// TIA Portal project "Yapisal Programlama" (V18)

(* hardware
DEVICE "S7-1200 station_1"  S7-1200 Station
   slot 0: "Rack_0"  S7-1200 Rack  Rack  V1.0
   slot 1: "PLC_1"  CPU 1214C DC/DC/Rly  6ES7 214-1HG40-0XB0  V4.6
*)

// ===== PLC "PLC_1"  CPU 1214C DC/DC/Rly =====

VAR_GLOBAL   // PLC tag table "Default tag table"
   "Start Butonu" AT %I0.0 : Bool;
   "Acil Stop Butonu" AT %I0.1 : Bool;
   "Reset Butonu" AT %I0.2 : Bool;
   "Yukarı Sensörü" AT %I0.3 : Bool;
   "Aşağı Sensörü" AT %I0.4 : Bool;
   "Piston Yukarı" AT %Q0.0 : Bool;
   "Piston Aşağı" AT %Q0.1 : Bool;
   "Sistem Start Mem" AT %M10.0 : Bool;
END_VAR

// folder: System blocks/Program resources

DATA_BLOCK "Counter 1"   // DB1
{ S7_Optimized_Access := 'TRUE' }
AUTHOR : Simatic
FAMILY : IEC
NAME : CNTR
VERSION : 1.0
// stored: InstanceOfName IEC_COUNTER
"IEC_COUNTER"
BEGIN
END_DATA_BLOCK

DATA_BLOCK "TIMER -1"   // DB2
{ S7_Optimized_Access := 'TRUE' }
AUTHOR : Simatic
FAMILY : IEC
NAME : IEC_TMR
VERSION : 1.0
// stored: InstanceOfName IEC_TIMER
"IEC_TIMER"
BEGIN
END_DATA_BLOCK

// folder: (top level)

FUNCTION "Normal Calisma" : Void   // FC1, LAD
{ S7_Optimized_Access := 'TRUE' }
VERSION : 0.1
BEGIN

REGION Network 1: SİSTEMİN BAŞLATILMASI
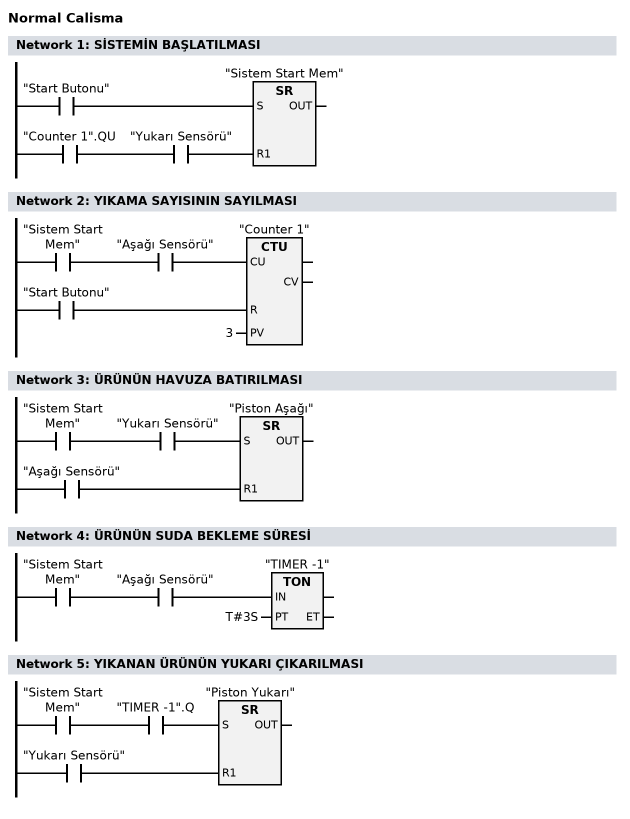
   RUNG wire#powerrail
      Contact( "Start Butonu" )
      S_SR(operand := "Sistem Start Mem", r1 := wire#w1)
   END_RUNG
   RUNG wire#powerrail
      Contact( "Counter 1".QU )
      Contact( "Yukarı Sensörü" )
   END_RUNG wire#w1
   // the same network as SCL:
   IF "Start Butonu" THEN
       "Sistem Start Mem" := TRUE;   // SR flip-flop
   END_IF;
   IF "Counter 1".QU AND "Yukarı Sensörü" THEN "Sistem Start Mem" := FALSE; END_IF;
END_REGION

REGION Network 2: YIKAMA SAYISININ SAYILMASI
   "Counter 1".CTU(CU := "Sistem Start Mem" AND "Aşağı Sensörü", R := "Start Butonu", PV := 3);
END_REGION

REGION Network 3: ÜRÜNÜN HAVUZA BATIRILMASI
   RUNG wire#powerrail
      Contact( "Sistem Start Mem" )
      Contact( "Yukarı Sensörü" )
      S_SR(operand := "Piston Aşağı", r1 := wire#w1)
   END_RUNG
   RUNG wire#powerrail
      Contact( "Aşağı Sensörü" )
   END_RUNG wire#w1
   // the same network as SCL:
   IF "Sistem Start Mem" AND "Yukarı Sensörü" THEN
       "Piston Aşağı" := TRUE;   // SR flip-flop
   END_IF;
   IF "Aşağı Sensörü" THEN "Piston Aşağı" := FALSE; END_IF;
END_REGION

REGION Network 4: ÜRÜNÜN SUDA BEKLEME SÜRESİ
   "TIMER -1".TON(IN := "Sistem Start Mem" AND "Aşağı Sensörü", PT := T#3S);
END_REGION

REGION Network 5: YIKANAN ÜRÜNÜN YUKARI ÇIKARILMASI
   RUNG wire#powerrail
      Contact( "Sistem Start Mem" )
      Contact( "TIMER -1".Q )
      S_SR(operand := "Piston Yukarı", r1 := wire#w1)
   END_RUNG
   RUNG wire#powerrail
      Contact( "Yukarı Sensörü" )
   END_RUNG wire#w1
   // the same network as SCL:
   IF "Sistem Start Mem" AND "TIMER -1".Q THEN
       "Piston Yukarı" := TRUE;   // SR flip-flop
   END_IF;
   IF "Yukarı Sensörü" THEN "Piston Yukarı" := FALSE; END_IF;
END_REGION
END_FUNCTION

FUNCTION "Acil Stop Calisma" : Void   // FC2, LAD
{ S7_Optimized_Access := 'TRUE' }
VERSION : 0.1
BEGIN

REGION Network 1: ACİL STOP BUTONUNA BASILDIĞINDA SİSTEMİN DURDURULMASI
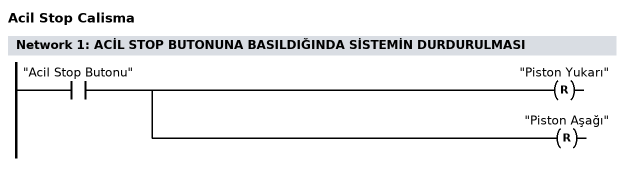
   RUNG wire#powerrail
      Contact( "Acil Stop Butonu" )
      wire#w1
      R_Coil( "Piston Yukarı" )
   END_RUNG
   RUNG wire#w1
      R_Coil( "Piston Aşağı" )
   END_RUNG
   // the same network as SCL:
   IF "Acil Stop Butonu" THEN
       "Piston Yukarı" := FALSE;
       "Piston Aşağı" := FALSE;
   END_IF;
END_REGION
END_FUNCTION

FUNCTION "Reset Calisma" : Void   // FC3, LAD
{ S7_Optimized_Access := 'TRUE' }
VERSION : 0.1
BEGIN

REGION Network 1: RESET BUTONUNA BASILDIĞINDA SİSTEMİN BAŞLANGIÇ KONUMUNA GETİRİLMESİ
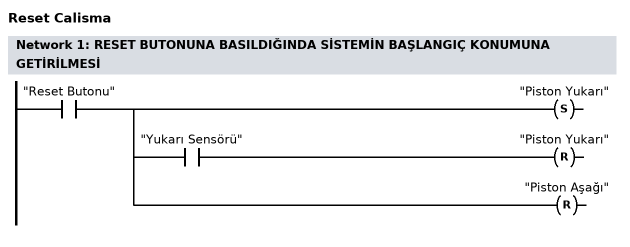
   RUNG wire#powerrail
      Contact( "Reset Butonu" )
      wire#w1
      S_Coil( "Piston Yukarı" )
   END_RUNG
   RUNG wire#w1
      Contact( "Yukarı Sensörü" )
      R_Coil( "Piston Yukarı" )
   END_RUNG
   RUNG wire#w1
      R_Coil( "Piston Aşağı" )
   END_RUNG
   // the same network as SCL:
   IF "Reset Butonu" THEN "Piston Yukarı" := TRUE; END_IF;
   IF "Reset Butonu" AND "Yukarı Sensörü" THEN "Piston Yukarı" := FALSE; END_IF;
   IF "Reset Butonu" THEN "Piston Aşağı" := FALSE; END_IF;
END_REGION
END_FUNCTION

ORGANIZATION_BLOCK "Ana Program"   // OB1, LAD, ProgramCycle
TITLE = "Main Program Sweep (Cycle)"
{ S7_Optimized_Access := 'TRUE' }
VERSION : 0.1
   VAR_INPUT
      Initial_Call : Bool;   // Initial call of this OB
      Remanence : Bool;   // =True, if remanent data are available
   END_VAR
BEGIN

REGION Network 1: ACİL STOP PROGRAMININ ÇAĞRILMASI
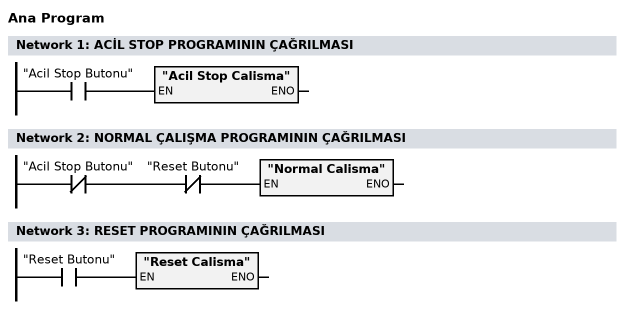
   RUNG wire#powerrail
      Contact( "Acil Stop Butonu" )
      "Acil Stop Calisma"()
   END_RUNG
   // the same network as SCL:
   IF "Acil Stop Butonu" THEN "Acil Stop Calisma"(); END_IF;
END_REGION

REGION Network 2: NORMAL ÇALIŞMA PROGRAMININ ÇAĞRILMASI
   RUNG wire#powerrail
      I_Contact( "Acil Stop Butonu" )
      I_Contact( "Reset Butonu" )
      "Normal Calisma"()
   END_RUNG
   // the same network as SCL:
   IF NOT "Acil Stop Butonu" AND NOT "Reset Butonu" THEN "Normal Calisma"(); END_IF;
END_REGION

REGION Network 3: RESET PROGRAMININ ÇAĞRILMASI
   RUNG wire#powerrail
      Contact( "Reset Butonu" )
      "Reset Calisma"()
   END_RUNG
   // the same network as SCL:
   IF "Reset Butonu" THEN "Reset Calisma"(); END_IF;
END_REGION
END_ORGANIZATION_BLOCK